// TIA Portal project "Task1_V18" (V18)

(* hardware
DEVICE "S7-1200 station_1"  S7-1200 Station
   slot 0: "Rack_0"  Rack  V1.0
   slot 1: "PLC_1"  CPU 1212C AC/DC/Rly  6ES7 212-1BE40-0XB0  V4.1
DEVICE "GSD device_1"  GSD.Device.PN
   slot 0: "Rack"  Rail  V1.0
   slot 0: "AL1100"  AL1100
   slot 1: "4 Ports_1"  AL1100
DEVICE "HMI_1"  TP700 Comfort
   slot 0: "HMI_1"  TP700 Comfort  6AV2 124-0GC01-0AX0  15.0.0.0
   slot 1: "HMI_RT_3"  TP700 Comfort  6AV2 124-0GC01-0AX0  15.0.0.0
   slot 5: "HMI_1.IE_CP_1"  PROFINET Interface  15.0.0.0
      slot 1: "PROFINET Schnittstelle_1"  PROFINET Interface
         slot 1: "Port_1"  Port
         slot 2: "Port_2"  Port
   slot 7: "HMI_1.MPI/DP_CP_1"  MPI/DP Interface  15.0.0.0
*)

// ===== PLC "PLC_1"  CPU 1212C AC/DC/Rly =====

VAR_GLOBAL   // PLC tag table "Default tag table"
   "Tag_1" AT %Q0.0 : Bool;
   "Tag_2" AT %M0.0 : Bool;
   "System_Byte" AT %MB1 : Byte;
   "FirstScan" AT %M1.0 : Bool;
   "DiagStatusUpdate" AT %M1.1 : Bool;
   "AlwaysTRUE" AT %M1.2 : Bool;
   "AlwaysFALSE" AT %M1.3 : Bool;
   "Clock_Byte" AT %MB0 : Byte;
   "Clock_5Hz" AT %M0.1 : Bool;
   "Clock_2.5Hz" AT %M0.2 : Bool;
   "Clock_2Hz" AT %M0.3 : Bool;
   "Clock_1.25Hz" AT %M0.4 : Bool;
   "Clock_1Hz" AT %M0.5 : Bool;
   "Clock_0.625Hz" AT %M0.6 : Bool;
   "Clock_0.5Hz" AT %M0.7 : Bool;
   "Tag_3" AT %M10.0 : Bool;
END_VAR

VAR_GLOBAL   // PLC tag table "RFID"
   "i_command_value" AT %IB90 : Byte;
   "i_command_ack" AT %I91.0 : Bool;
   "i_command_end" AT %I91.1 : Bool;
   "i_tag_present" AT %I91.2 : Bool;
   "i_antenna_deactivated" AT %I91.3 : Bool;
   "i_read_value_0" AT %IW92 : Int;
   "i_read_value_1" AT %IW94 : Int;
   "i_read_value_2" AT %IW96 : Int;
   "i_read_value_3" AT %IW98 : Int;
   "q_command_value" AT %QB84 : Byte;
   "q_start_r/w" AT %Q85.0 : Bool;
   "q_antenna_deactivate" AT %Q85.3 : Bool;
   "q_write_value_0" AT %QW86 : Int;
   "q_write_value_1" AT %QW88 : Int;
   "q_write_value_2" AT %QW90 : Int;
   "q_write_value_3" AT %QW92 : Int;
END_VAR

TYPE "RFID_IOLink"
VERSION : 0.1
   STRUCT
      Input : Struct
         command_ack : Bool;
         command_end : Bool;
         tag_present : Bool;
         Antenna_deactivated : Bool;
         command_value : Byte;
         read_values : Array[0..3] of Int;
      END_STRUCT;
      Output : Struct
         "Start_r/w" : Bool;
         Deactivate_antenna : Bool;
         command_value : Byte;   // 0= read UID, 1=Auto-read, 2=Auto-write, 3=read, 4=write
         write_values : Array[0..3] of Int;
      END_STRUCT;
   END_STRUCT;
END_TYPE

DATA_BLOCK "ModeInterface"   // DB2
{ S7_Optimized_Access := 'TRUE' }
VERSION : 0.1
   VAR
      AssignSupervisor : Bool;
      AssignService : Bool;
      AssignOperator : Bool;
      TagDisable : Bool;
      WriteID : Bool;
      "ActuateQ0.0" : Bool;
      LoginStatus : Int;
      SetTimeDelay : Time;
      CurrentTimeDelay : Time;
   END_VAR
BEGIN
END_DATA_BLOCK

// folder: Login

DATA_BLOCK "Login_logic_DB"   // DB13
{ S7_Optimized_Access := 'TRUE' }
VERSION : 0.1
// stored: InstanceOfName Login_logic
"Login_logic"
BEGIN
END_DATA_BLOCK

// folder: RFID

DATA_BLOCK "RFIDData"   // DB1
{ S7_Optimized_Access := 'FALSE' }
VERSION : 0.1
   VAR
      RFID : "RFID_IOLink";
   END_VAR
BEGIN
   RFID.Output.command_value := 16#1;
END_DATA_BLOCK

// folder: System blocks/Program resources

DATA_BLOCK "IEC_Timer_0_DB"   // DB3
{ S7_Optimized_Access := 'TRUE' }
AUTHOR : Simatic
FAMILY : IEC
NAME : IEC_TMR
VERSION : 1.0
// stored: InstanceOfName IEC_TIMER
"IEC_TIMER"
BEGIN
END_DATA_BLOCK

// folder: (top level)

ORGANIZATION_BLOCK "Main"   // OB1, LAD, ProgramCycle
TITLE = "Main Program Sweep (Cycle)"
{ S7_Optimized_Access := 'TRUE' }
VERSION : 0.1
   VAR_INPUT
      Initial_Call : Bool;   // Initial call of this OB
      Remanence : Bool;   // =True, if remanent data are available
   END_VAR
BEGIN

REGION Network 1: Read values from RFID
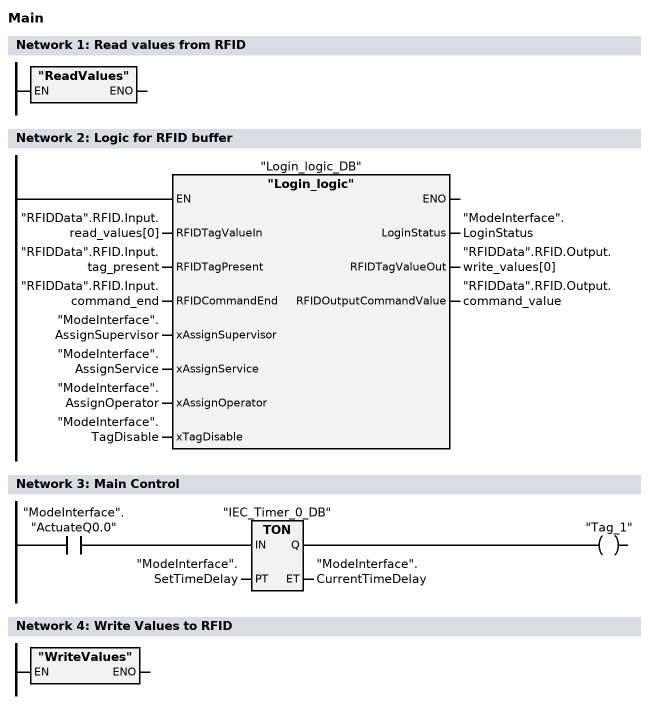
   RUNG wire#powerrail
      "ReadValues"()
   END_RUNG
   // the same network as SCL:
   "ReadValues"();
END_REGION

REGION Network 2: Logic for RFID buffer
   RUNG wire#powerrail
      "Login_logic_DB"(RFIDTagValueIn := "RFIDData".RFID.Input.read_values[0], RFIDTagPresent := "RFIDData".RFID.Input.tag_present, RFIDCommandEnd := "RFIDData".RFID.Input.command_end, xAssignSupervisor := "ModeInterface".AssignSupervisor, xAssignService := "ModeInterface".AssignService, xAssignOperator := "ModeInterface".AssignOperator, xTagDisable := "ModeInterface".TagDisable, LoginStatus => "ModeInterface".LoginStatus, RFIDTagValueOut => "RFIDData".RFID.Output.write_values[0], RFIDOutputCommandValue => "RFIDData".RFID.Output.command_value)
   END_RUNG
   // the same network as SCL:
   "Login_logic_DB"(RFIDTagValueIn := "RFIDData".RFID.Input.read_values[0],   // "Login_logic"
                    RFIDTagPresent := "RFIDData".RFID.Input.tag_present,
                    RFIDCommandEnd := "RFIDData".RFID.Input.command_end,
                    xAssignSupervisor := "ModeInterface".AssignSupervisor,
                    xAssignService := "ModeInterface".AssignService,
                    xAssignOperator := "ModeInterface".AssignOperator,
                    xTagDisable := "ModeInterface".TagDisable,
                    LoginStatus => "ModeInterface".LoginStatus,
                    RFIDTagValueOut => "RFIDData".RFID.Output.write_values[0],
                    RFIDOutputCommandValue => "RFIDData".RFID.Output.command_value);
END_REGION

REGION Network 3: Main Control
   "IEC_Timer_0_DB".TON(IN := "ModeInterface"."ActuateQ0.0",
                        PT := "ModeInterface".SetTimeDelay,
                        ET => "ModeInterface".CurrentTimeDelay);
   "Tag_1" := "IEC_Timer_0_DB".Q;
END_REGION

REGION Network 4: Write Values to RFID
   RUNG wire#powerrail
      "WriteValues"()
   END_RUNG
   // the same network as SCL:
   "WriteValues"();
END_REGION
END_ORGANIZATION_BLOCK

// folder: Login

FUNCTION_BLOCK "Login_logic"   // FB8, FBD
TITLE = Tag Management
{ S7_Optimized_Access := 'TRUE' }
VERSION : 0.1
   VAR_INPUT
      RFIDTagValueIn : Int;
      RFIDTagPresent : Bool;
      RFIDCommandEnd : Bool;
   END_VAR
   VAR_OUTPUT
      LoginStatus : Int;
      RFIDTagValueOut : Int;
      RFIDOutputCommandValue : Int;
   END_VAR
   VAR_IN_OUT
      xAssignSupervisor : Bool;
      xAssignService : Bool;
      xAssignOperator : Bool;
      xTagDisable : Bool;
   END_VAR
   VAR
      tonTagPresent : TON_TIME;
      Flag : Bool;
   END_VAR
   VAR_TEMP   // added for the SCL form of the ladder/FBD networks
      _w1 : Bool;
   END_VAR
BEGIN

REGION Network 1: Login supervisor / Supervisor Login function
   // RFID Value 5801 represents Supervisor with login status 2
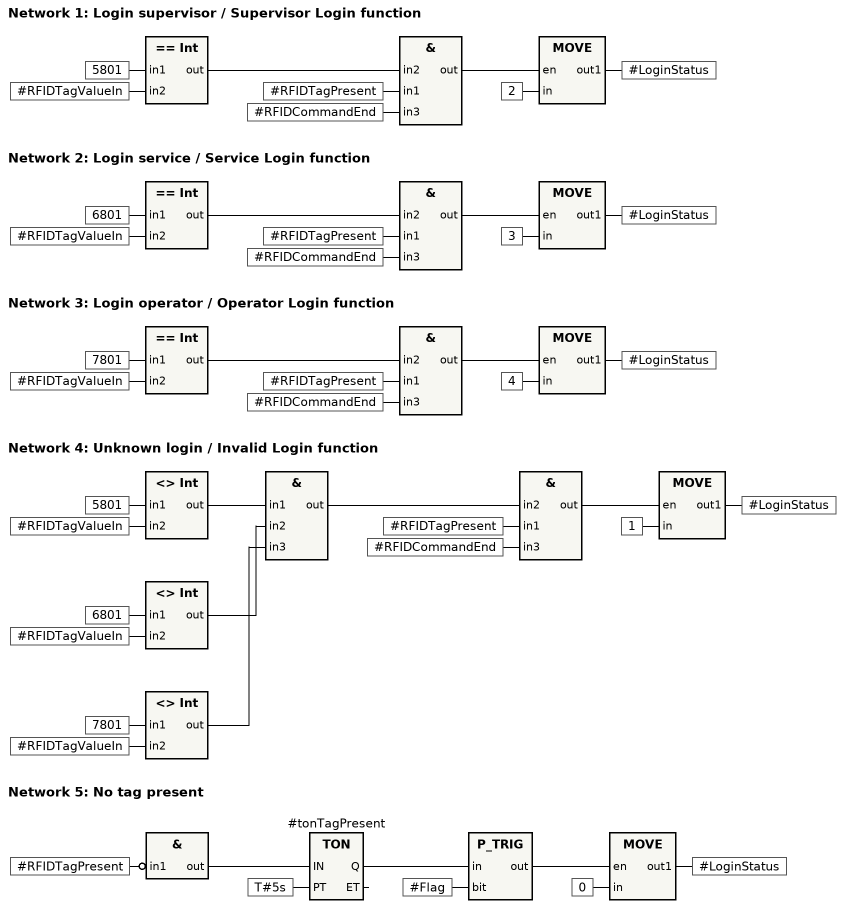
   IF (5801 = #RFIDTagValueIn) AND #RFIDTagPresent AND #RFIDCommandEnd THEN #LoginStatus := 2; END_IF;
END_REGION

REGION Network 2: Login service / Service Login function
   // RFID Value 6801 represents Service with login status 3
   IF (6801 = #RFIDTagValueIn) AND #RFIDTagPresent AND #RFIDCommandEnd THEN #LoginStatus := 3; END_IF;
END_REGION

REGION Network 3: Login operator / Operator Login function
   // RFID Value 7801 represents Operator with login status 4
   IF (7801 = #RFIDTagValueIn) AND #RFIDTagPresent AND #RFIDCommandEnd THEN #LoginStatus := 4; END_IF;
END_REGION

REGION Network 4: Unknown login / Invalid Login function
   // with login status 1
   IF (5801 <> #RFIDTagValueIn) AND (6801 <> #RFIDTagValueIn) AND (7801 <> #RFIDTagValueIn) AND #RFIDTagPresent AND #RFIDCommandEnd THEN
       #LoginStatus := 1;
   END_IF;
END_REGION

REGION Network 5: No tag present
   // with login status 0
   #tonTagPresent(IN := NOT #RFIDTagPresent, PT := T#5s);   // TON
   #_w1 := #tonTagPresent.Q AND NOT #Flag;   // rising edge
   #Flag := #tonTagPresent.Q;
   IF #_w1 THEN #LoginStatus := 0; END_IF;
END_REGION

REGION Network 6: Tag Managment / Tag Management
   // Command value 2 = Automatic write and Command value 1 = Automatic read
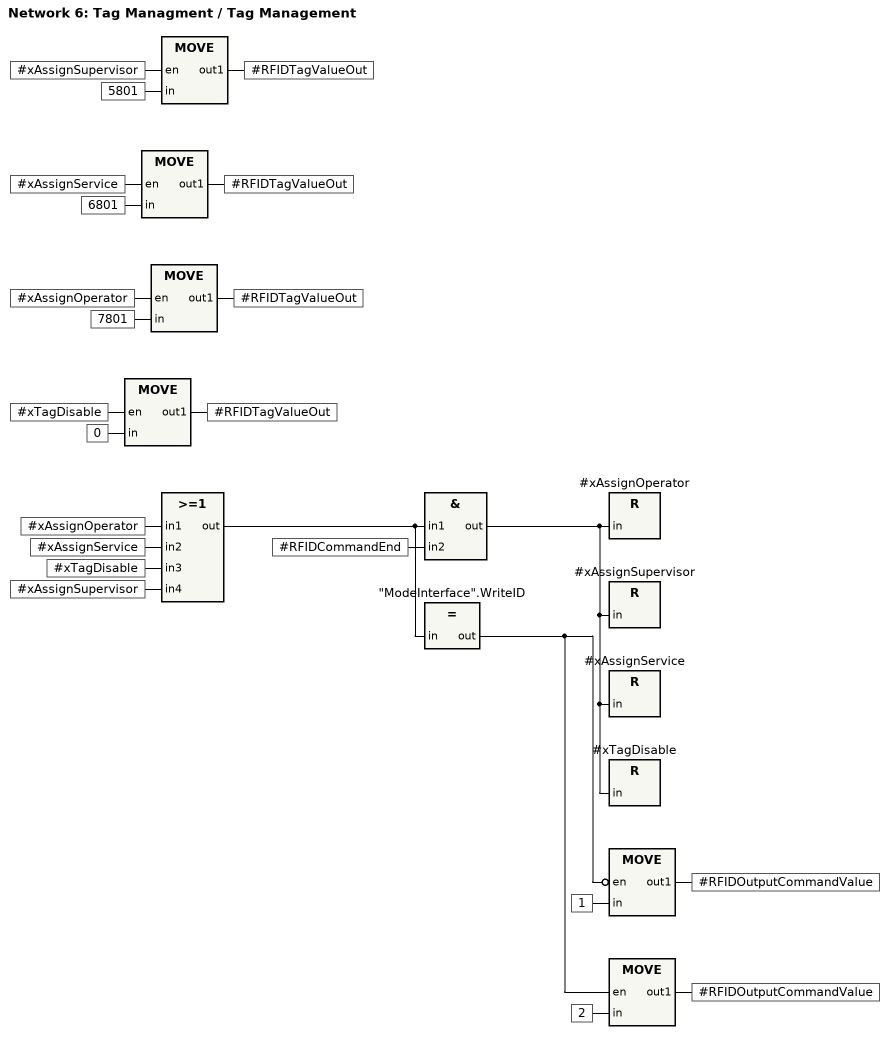
   IF #xAssignSupervisor THEN #RFIDTagValueOut := 5801; END_IF;
   IF #xAssignService THEN #RFIDTagValueOut := 6801; END_IF;
   IF #xAssignOperator THEN #RFIDTagValueOut := 7801; END_IF;
   IF #xTagDisable THEN #RFIDTagValueOut := 0; END_IF;
   #_w1 := #xAssignOperator OR #xAssignService OR #xTagDisable OR #xAssignSupervisor;
   IF #_w1 AND #RFIDCommandEnd THEN
       #xAssignOperator := FALSE;
       #xAssignSupervisor := FALSE;
       #xAssignService := FALSE;
       #xTagDisable := FALSE;
   END_IF;
   "ModeInterface".WriteID := #_w1;
   IF NOT #_w1 THEN #RFIDOutputCommandValue := 1; END_IF;
   IF #_w1 THEN #RFIDOutputCommandValue := 2; END_IF;
END_REGION
END_FUNCTION_BLOCK

// folder: RFID

FUNCTION "ReadValues" : Void   // FC1, SCL
{ S7_Optimized_Access := 'TRUE' }
VERSION : 0.1
BEGIN
   //Reading value from RFID
   "RFIDData".RFID.Input.command_ack:="i_command_ack";
   "RFIDData".RFID.Input.command_value:="i_command_value";
   "RFIDData".RFID.Input.command_end:="i_command_end";
   "RFIDData".RFID.Input.tag_present:="i_tag_present";
   "RFIDData".RFID.Input.Antenna_deactivated:="i_antenna_deactivated";
   "RFIDData".RFID.Input.read_values[0]:="i_read_value_0";
   "RFIDData".RFID.Input.read_values[1]:="i_read_value_1";
   "RFIDData".RFID.Input.read_values[2]:="i_read_value_2";
   "RFIDData".RFID.Input.read_values[3]:="i_read_value_3";
END_FUNCTION

FUNCTION "WriteValues" : Void   // FC2, SCL
{ S7_Optimized_Access := 'TRUE' }
VERSION : 0.1
BEGIN
   //Writing values to RFID
   "q_command_value" := "RFIDData".RFID.Output.command_value;
   "q_start_r/w" := "RFIDData".RFID.Output."Start_r/w";
   "q_antenna_deactivate" := "RFIDData".RFID.Output.Deactivate_antenna;
   "q_write_value_0" := "RFIDData".RFID.Output.write_values[0];
   "q_write_value_1" := "RFIDData".RFID.Output.write_values[1];
   "q_write_value_2" := "RFIDData".RFID.Output.write_values[2];
   "q_write_value_3" := "RFIDData".RFID.Output.write_values[3];
END_FUNCTION

(* ===== HMI "HMI_RT_3" =====
system functions are stored by id; their names below are inferred from use
connection "HMI_Connection_1": ETHERNET, S7_1200_OMS

HMI tags "Standard-Variablentabelle"
   "ActuatuteQ0.0" : Bool = PLC ModeInterface."ActuateQ0.0" AT %DB1.DBX0.0, 100 ms
   "SetDelayQ0.0" : Time = PLC ModeInterface.SetTimeDelay AT %DB1.DBD0, 100 ms
   "CurrentDelayQ0.0" : Time = PLC ModeInterface.CurrentTimeDelay AT %DB1.DBD0, 100 ms
   "FeedbackQ0.0" : Bool = PLC Tag_1 AT %Q0.0, 100 ms

HMI tags "Login"
   "password" : WString[254], internal
   "Login" : WString[254], internal
   "RFID_Tag_present" : Bool = PLC RFIDData.RFID.Input.tag_present AT %DB1.DBX0.2, 100 ms
   "xAssignSupervisor" : Bool = PLC ModeInterface.AssignSupervisor AT %DB1.DBX0.0, 100 ms
   "xRFIDValue" : Int = PLC RFIDData.RFID.Input.read_values[0] AT %DB1.DBW2, 100 ms
   "xAssignOperator" : Bool = PLC ModeInterface.AssignOperator AT %DB1.DBX0.0, 100 ms
   "xAssignService" : Bool = PLC ModeInterface.AssignService AT %DB1.DBX0.0, 100 ms
   "xDisableTag" : Bool = PLC ModeInterface.TagDisable AT %DB1.DBX0.0, 100 ms
   "status_login" : Int = PLC ModeInterface.LoginStatus AT %DB1.DBW0, 100 ms
      on ChangeValue: "VBFunction_2"()
   "getuser" : WString[254], internal
   "getuser_1" : WString[254], internal
   "1Hz" : Bool = PLC Clock_1Hz AT %M0.5, 500 ms
      on ChangeValue: "VBFunction_1"(); function_f41c6f6c("getuser")

discrete alarms
   2: 'Timeout extend Drawer Magazin 1', class Magazin 1, trigger "Errors_wErrorsMagazine1" bit 1
   19: 'Slide 1 full, please empty Slide 1 and confirm', class Slides, trigger "Errors_wErrorsSlides" bit 1
   23: 'Pressure failure, plese adjust pressure level', class System Error, trigger "Errors_wSystem" bit 1
   10: 'Timeout extend Cylinder 1', class Sorting Unit, trigger "Errors_wErrorsSortingUnit" bit 1
   21: 'Slide 3 full, please empty Slide 3 and confirm', class Slides, trigger "Errors_wErrorsSlides" bit 3
   17: 'No RFID-Tag detected, please check workpiece', class Sorting Unit, trigger "Errors_wErrorsSortingUnit" bit 8
   14: 'Timeout extend Cylinder 3', class Sorting Unit, trigger "Errors_wErrorsSortingUnit" bit 5
   4: 'No Workpiece detected, check belt conveyor and Magazine 2', class Magazin 1, trigger "Errors_wErrorsMagazine1" bit 3
   8: 'No Workpiece detected, check belt conveyor and Magazine 2', class Magazin 2, trigger "Errors_wErrorsMagazine2" bit 3
   11: 'Timeout retract Cylinder 1', class Sorting Unit, trigger "Errors_wErrorsSortingUnit" bit 2
   7: 'Timeout retract Drawer Magazin 2', class Magazin 2, trigger "Errors_wErrorsMagazine2" bit 2
   13: 'Timeout retract Cylinder 2', class Sorting Unit, trigger "Errors_wErrorsSortingUnit" bit 4
   12: 'Timeout extend Cylinder 2', class Sorting Unit, trigger "Errors_wErrorsSortingUnit" bit 3
   15: 'Timeout retract Cylinder 3', class Sorting Unit, trigger "Errors_wErrorsSortingUnit" bit 6
   16: 'Workpiece missing, pleace check magazines and belt conveyor', class Sorting Unit, trigger "Errors_wErrorsSortingUnit" bit 7
   6: 'Timeout extend Drawer Magazin 2', class Magazin 2, trigger "Errors_wErrorsMagazine2" bit 1
   3: 'Timeout retract Drawer Magazin 1', class Magazin 1, trigger "Errors_wErrorsMagazine1" bit 2
   20: 'Slide 2 full, please empty Slide 2 and confirm', class Slides, trigger "Errors_wErrorsSlides" bit 2
   26: 'Workpiece could not be sorted out, please empty Slide 3 and confirm', class Slides, trigger "Errors_wErrorsSlides" bit 6
   25: 'Workpiece could not be sorted out, please empty Slide 2 and confirm', class Slides, trigger "Errors_wErrorsSlides" bit 5
   24: 'Workpiece could not be sorted out, please empty Slide 1 and confirm', class Slides, trigger "Errors_wErrorsSlides" bit 4
   22: 'Emergency Stop activ, please check EM-Stop button and reset', class System Error, trigger "Errors_wSystem" bit 0

text list "User Administration": 0..5800 'Not Used / Please scan valid tag'; 5801 'Supervisor'; 6801 'Service'; 7801 'Operator'

screen "Main" 800x426, template "Vorlage_1"
   GraphicView "Grafikanzeige_1" at 552,113 size 105x120; Picture "RFID Tag"
   Button "Schaltfläche_2" at 529,240 size 155x36; TextOff 'Tag Management Tag Management'; Authorization "TagManagement"
      on Press: ActivateScreen("Tag Management", 0)
   Button "Schaltfläche_1" at 558,116 size 97x116; TextOff 'Text'
      on Press: ActivateScreen("Tag Management", 0)
   IOField "I/O field_1" at 154,118 size 96x32; FormatPattern ????????????
      ProcessValue <- "Login"
   IOField "I/O field_2" at 340,118 size 96x32; FormatPattern ????????????????????????????????????????????????????????????????????????????????
      ProcessValue <- "password"
   TextField "Text field_2" at 122,123 size 24x23; Text 'Id / ID'
   TextField "Text field_3" at 254,122 size 91x23; Text 'Password'
   TextField "Text field_4" at 143,78 size 282x27; Text 'Kindly scan your ID to Login'
      Visibility <- "status_login"
   TextField "Text field_6" at 172,65 size 231x50; Text 'Authorized access! Click on Login button'
      Visibility <- "status_login"
   TextField "Text field_5" at 172,78 size 235x27; Text 'Unauthorized access !'
      Visibility <- "status_login"
   Button "Button_3" at 282,161 size 96x39; TextOff 'Log out / Logout'
      on Press: function_f23ef4c9(); "VBFunction_2"()
   UserView "User view_1" at 69,213 size 404x158
   TextField "Text field_1" at 278,5 size 253x32; Text 'User Login via RFID'
   Button "Schaltfläche_4" at 531,282 size 153x32; TextOff 'Parameters'; Authorization "Parameters"
      on Click: function_efd93a16("Parameter", 275, 75, -1, -1, 1)
   Button "Schaltfläche_7" at 531,322 size 152x38; TextOff 'Reverse / Actuate Q0.0'; Authorization "Actuate"
      on Press: function_b14e0dd5("ActuatuteQ0.0", 0)
      Appearance <- "FeedbackQ0.0"
   Button "Button_1" at 168,163 size 102x36; TextOff 'Login'
      on Press: function_a9b89908("password", "Login")
   Bar "Bar_1" at 688,323 size 104x36; MinimumValue 0; MaximumValue 100
      MaximumValue <- "SetDelayQ0.0"
      ProcessValue <- "CurrentDelayQ0.0"
   IOField "I/O field_3" at 687,367 size 107x28; FormatPattern s9999
      ProcessValue <- "SetDelayQ0.0"
   TextField "Text field_7" at 493,372 size 211x23; Text 'Set Time delay (in ms)'

screen "Tag Management" 800x426
   TextField "Textfeld_1" at 156,109 size 187x23; Text 'Check Status of Tag'
   TextField "Textfeld_12" at 76,-22 size 45x29; Text 'Tag Management'
   Rectangle "Rectangle_1" at 334,111 size 17x18
      Appearance <- "RFID_Tag_present"
   TextField "Textfeld_2" at 354,109 size 114x23; Text 'Tag present'
   TextField "Textfeld_3" at 203,156 size 48x23; Text 'Task'
   TextField "Textfeld_5" at 329,156 size 101x23; Text 'Supervisor'
   TextField "Textfeld_6" at 429,156 size 71x23; Text 'Service'
   TextField "Textfeld_7" at 506,156 size 86x23; Text 'Operator'
   TextField "Textfeld_8" at 591,156 size 57x23; Text 'Guest'
   TextField "Textfeld_9" at 201,184 size 121x42; Text 'Tag Management'
   TextField "Textfeld_10" at 201,239 size 102x42; Text 'Parameter Change'
   TextField "Textfeld_11" at 201,299 size 102x42; Text 'Operation Control'
   TextField "Textfeld_14" at 201,357 size 103x42; Text 'Monitor/ Navigation'
   Switch "Switch_1" at 283,50 size 98x47; TextOn 'Assign Supervisor'; CaptionText 'Switch'; TextOff 'Assign Supervisor'
      ProcessValue <- "xAssignSupervisor"
      Appearance <- "xAssignSupervisor"
   Switch "Switch_2" at 393,50 size 77x47; TextOn 'Assign Service'; CaptionText 'Switch'; TextOff 'Assign Service'
      ProcessValue <- "xAssignService"
      Appearance <- "xAssignService"
   Switch "Switch_3" at 480,50 size 88x47; TextOn 'Assign Operator'; CaptionText 'Switch'; TextOff 'Assign Operator'
      ProcessValue <- "xAssignOperator"
      Appearance <- "xAssignOperator"
   Switch "Switch_4" at 580,50 size 77x47; TextOn 'Disable Tag'; CaptionText 'Switch'; TextOff 'Disable Tag'
      ProcessValue <- "xDisableTag"
      Appearance <- "xDisableTag"
   Group "Group" at 356,198 size 27x19
   Group "Group_1" at 358,252 size 27x19
   Group "Group_2" at 357,309 size 27x19
   Group "Group_4" at 357,373 size 27x19
   Group "Group_5" at 451,252 size 27x19
   Group "Group_6" at 450,309 size 27x19
   Group "Group_8" at 450,373 size 27x19
   Group "Group_9" at 530,310 size 27x19
   Group "Group_11" at 530,374 size 27x19
   Group "Group_12" at 602,373 size 27x19
   TextField "Textfeld_15" at 153,53 size 110x42; Text 'Select Tag Assignment Select Tag Assignment'
   TextField "Text field_1" at 301,10 size 221x32; Text 'Tag Management'
   Button "Schaltfläche_2" at 13,381 size 80x36; TextOff 'Tag Management Back'; Authorization "TagManagement"
      on Press: ActivateScreen("Main", 0)
   SymbolicIOField "Symbolic I/O field_1" at 461,107 size 196x32; TextOff '0'; TextOn '1'; TextList "User Administration"
      ProcessValue <- "xRFIDValue"

PopupScreen "Parameter" 240x300
   TextField "Textfeld_12" at 6,2 size 111x29; Text 'Belt Conveyor / Parameters'
   Button "Schaltfläche_1" at 205,2 size 32x32; TextOff 'X / x'
      on Click: function_efd93a16("Parameter", 0, 0, -1, -1, 1)
   Button "Schaltfläche_3" at 0,260 size 240x40; TextOff 'Close'
      on Click: function_efd93a16("Parameter", 0, 0, -1, -1, 1)
   IOField "I/O field_1" at 87,121 size 73x32; FormatPattern s99999
      ProcessValue <- "SetDelayQ0.0"
   TextField "Text field_1" at 45,69 size 178x23; Text 'Q0.0 On delay time'
   TextField "Text field_2" at 91,92 size 69x23; Text '(in ms)'

VB script "VBFunction_2"
   'Tip:
   ' 1. Use the <CTRL+SPACE> or <CTRL+I> shortcut to open a list of all objects and functions
   ' 2. Write the code using the HMI Runtime object.
   '  Example: HmiRuntime.Screens("Screen_1").
   ' 3. Use the <CTRL+J> shortcut to create an object reference.
   'Write the code as of this position:
   
   'If user press logout button, user and password field should be empty
   
   SmartTags("Login") = ""
   SmartTags("password") = ""

VB script "VBFunction_1"
   'Tip:
   ' 1. Use the <CTRL+SPACE> or <CTRL+I> shortcut to open a list of all objects and functions
   ' 2. Write the code using the HMI Runtime object.
   '  Example: HmiRuntime.Screens("Screen_1").
   ' 3. Use the <CTRL+J> shortcut to create an object reference.
   'Write the code as of this position:
   
   'Status Login = 0 it means no user is logged in or no tag is present
   
   If SmartTags("status_login") = 0 Then
   	SmartTags("Login") = ""
   	SmartTags("password") = ""
   End If
   
   
   'Status Login = 1 it means invalid user or unauthorized access
   
   If SmartTags("status_login") = 1 Then
   	SmartTags("Login") = "xxxx"
   	SmartTags("password") = "xxxx"
   End If
   
   'Status Login = 2 it means Supervisor is logged in
   
   If SmartTags("status_login") = 2 Then
   	SmartTags("Login") = "Supervisor"
   	SmartTags("password") = "c5801"
   End If
   
   
   'Status Login = 3 it means Service is logged in
   
   If SmartTags("status_login") = 3 Then
   	SmartTags("Login") = "Service"
   	SmartTags("password") = "c6801"
   End If
   
   'Status Login = 4 it means Operator is logged in
   
   If SmartTags("status_login") = 4 Then
   	SmartTags("Login") = "Operator"
   	SmartTags("password") = "c7801"
   End If
   
   'Fucntion to display the name of user in top right screen
   Dim length
   length = Len (SmartTags("getuser"))
   If length < 1 Then
   	SmartTags("getuser_1") = "Guest"
   Else
   	SmartTags("getuser_1") = SmartTags("getuser")
   End if
*)